Fanuc KAREL source: KX00025.KL

PROGRAM KX00025
%NOLOCKGROUP
%COMMENT = 'Feature sample'
VAR
  I: INTEGER
  J: INTEGER
  B: BOOLEAN
  F: FILE
  S: STRING[80]
  P: XYZWPR
BEGIN
  I = 1
END KX00025
